FUNCTION FC 1 : VOID
BEGIN
NETWORK
      A MW 10
END_FUNCTION
